Fanuc KAREL source: kb00033.KL

-- PROVISIONAL review KL for V940-1; original PC SHA256 4d0a96df51ffc5bf11c0d813cc1215c8df090be07bdfdd10ec53915a7ef05a94
-- Incomplete behavior may be omitted. Consult companion uncertainty JSON. Do not deploy.
PROGRAM KB00033
%NOLOCKGROUP
BEGIN
  -- V9_ZERO_TABLE_METADATA_HINT layout=0002_ascii; no indexed target words; source/name/runtime held
  -- UNRESOLVED_PC offsets 5-14; opcodes 3F,75
  -- UNRESOLVED_PC offsets 19-26; opcodes 9D,23
  -- UNRESOLVED_PC offsets 31-57; opcodes 27,22,22,2A,22,27,9D,31
  -- UNRESOLVED_PC offsets 62-66; opcodes 7F
END KB00033
